SUBAPPLICATION SubType
  (* Standard: 61499-1; Description: Copyright (c) 2026 Martin Erich Jobst This program and the accompanying materials are made available under the terms of the Eclipse Public License 2.0 which is available at https://www.eclipse.org/legal/epl-2.0/ SPDX-License-Identifier: EPL-2.0 *)
  (* Version 1.0, 2026-11-18, Martin Jobst *)
  PACKAGE lib::VarConfigInstance::support;
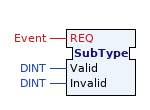
  EVENT_INPUT
    REQ;
  END_EVENT
  VAR_INPUT
    Valid : DINT;
    Invalid : DINT;
  END_VAR
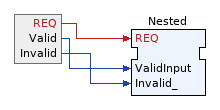
  SUBAPPLICATION Nested
    EVENT_INPUT
      REQ;
    END_EVENT
    VAR_INPUT
      ValidInput : DINT;
      Invalid_ : DINT;
    END_VAR
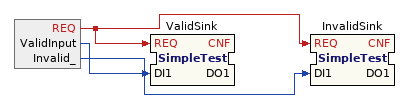
    FBS
      ValidSink : lib::VarConfigInstance::support::SimpleTest;
      InvalidSink : lib::VarConfigInstance::support::SimpleTest;
    END_FBS
    EVENT_CONNECTIONS
      REQ TO ValidSink.REQ;
      REQ TO InvalidSink.REQ;
    END_CONNECTIONS
    DATA_CONNECTIONS
      ValidInput TO ValidSink.DI1;
      Invalid_ TO InvalidSink.DI1;
    END_CONNECTIONS
  END_SUBAPPLICATION
  EVENT_CONNECTIONS
    REQ TO Nested.REQ;
  END_CONNECTIONS
  DATA_CONNECTIONS
    Valid TO Nested.ValidInput;
    Invalid TO Nested.Invalid_;
  END_CONNECTIONS
END_SUBAPPLICATION
